// Composition of the event services, built once in a composition root (see GVL_EventDefaults).
// The setters let an application swap a single service; set them before the first event is raised.
FUNCTION_BLOCK FB_EventContext IMPLEMENTS I_EventContext
VAR
	_ipTexts		: I_TextProvider;
	_ipLanguage		: I_LanguageProvider;
	_ipFormatter	: I_TextFormatter;
	_ipEventEntries	: I_EventEntryProvider;
END_VAR

METHOD FB_init : BOOL
VAR_INPUT
	bInitRetains	: BOOL;
	bInCopyCode		: BOOL;
	ipTexts			: I_TextProvider;
	ipLanguage		: I_LanguageProvider;
	ipFormatter		: I_TextFormatter;
	ipEventEntries	: I_EventEntryProvider;
END_VAR
_ipTexts := ipTexts;
_ipLanguage := ipLanguage;
_ipFormatter := ipFormatter;
_ipEventEntries := ipEventEntries;
END_METHOD

PROPERTY Texts : I_TextProvider
GET
Texts := _ipTexts;
END_GET
SET
_ipTexts := Texts;
END_SET
END_PROPERTY

PROPERTY Language : I_LanguageProvider
GET
Language := _ipLanguage;
END_GET
SET
_ipLanguage := Language;
END_SET
END_PROPERTY

PROPERTY Formatter : I_TextFormatter
GET
Formatter := _ipFormatter;
END_GET
SET
_ipFormatter := Formatter;
END_SET
END_PROPERTY

PROPERTY EventEntries : I_EventEntryProvider
GET
EventEntries := _ipEventEntries;
END_GET
SET
_ipEventEntries := EventEntries;
END_SET
END_PROPERTY

END_FUNCTION_BLOCK

(* stored: Version 1.1.0.1, ProductVersion 3.1.4026.26
   POU FB_EventContext: Id {d1caea09-763a-4400-95a8-32d8d88b23a9}, SpecialFunc None
   Method FB_init: Id {f6f1e899-e3f4-4807-968a-9a090c7898d9}
   Property Texts: Id {1c9ca600-785c-40c1-9b3e-5f97eb756a7e}
   Get Get: Id {af7b2781-f1ca-418e-8cc4-a8354c7d544d}
   Set Set: Id {d53de5c5-6a52-429e-881d-8c0d79a39c59}
   Property Language: Id {71f66701-5201-42a1-af3b-d49b1ab4f252}
   Get Get: Id {c7a437be-e62a-4a75-a806-fc71f1e69c8f}
   Set Set: Id {29851781-8028-4e4a-897c-a4dce799b889}
   Property Formatter: Id {7aa437eb-2ecf-412f-8fbf-0a1cde23722b}
   Get Get: Id {b4bee6bc-eefe-46fb-8874-49e70efa9fd3}
   Set Set: Id {a2b8511e-8bbe-441d-a293-61809fb1c441}
   Property EventEntries: Id {c81f2f39-765b-451b-9c4e-4a0ac4f0a59f}
   Get Get: Id {215c3038-be8a-4b06-8071-a1f0f33a4988}
   Set Set: Id {7ee7a522-1646-464c-9acb-8caa6b306e0e} *)
